// --- Siemens Structured Format ---
DATA_BLOCK "model__HS8_IW10_"
{ S7_Optimized_Access := 'TRUE' }
VERSION :
NON_RETAIN
   VAR
      W_i : ARRAY[0..7, 0..39] OF REAL;
      W_f : ARRAY[0..7, 0..39] OF REAL;
      W_g : ARRAY[0..7, 0..39] OF REAL;
      W_o : ARRAY[0..7, 0..39] OF REAL;
      R_i : ARRAY[0..7, 0..7] OF REAL;
      R_f : ARRAY[0..7, 0..7] OF REAL;
      R_g : ARRAY[0..7, 0..7] OF REAL;
      R_o : ARRAY[0..7, 0..7] OF REAL;
      B_i : ARRAY[0..7] OF REAL;
      B_f : ARRAY[0..7] OF REAL;
      B_g : ARRAY[0..7] OF REAL;
      B_o : ARRAY[0..7] OF REAL;
      FC_W : ARRAY[0..39, 0..7] OF REAL;
      FC_B : ARRAY[0..39] OF REAL;
   END_VAR
BEGIN

      W_i[0,0] := -0.07214709;
      W_i[0,1] := 0.05972328;
      W_i[0,2] := 0.02437277;
      W_i[0,3] := -0.07067372;
      W_i[0,4] := 0.15626091;
      W_i[0,5] := 0.03422371;
      W_i[0,6] := -0.01010964;
      W_i[0,7] := 0.24618091;
      W_i[0,8] := 0.19837169;
      W_i[0,9] := -0.16936609;
      W_i[0,10] := -0.03685989;
      W_i[0,11] := -0.34127542;
      W_i[0,12] := 0.16145179;
      W_i[0,13] := -0.03563828;
      W_i[0,14] := -0.03820900;
      W_i[0,15] := 0.03625023;
      W_i[0,16] := -0.00035658;
      W_i[0,17] := 0.05683306;
      W_i[0,18] := 0.01328012;
      W_i[0,19] := 0.01230632;
      W_i[0,20] := -0.02302203;
      W_i[0,21] := 0.29246566;
      W_i[0,22] := -0.40551317;
      W_i[0,23] := -0.00420093;
      W_i[0,24] := -0.49537772;
      W_i[0,25] := -0.37926760;
      W_i[0,26] := -0.32712772;
      W_i[0,27] := -0.47364110;
      W_i[0,28] := -0.02835605;
      W_i[0,29] := -0.19270489;
      W_i[0,30] := -0.02380528;
      W_i[0,31] := -0.25659311;
      W_i[0,32] := -0.07342248;
      W_i[0,33] := 0.12401358;
      W_i[0,34] := -0.00912032;
      W_i[0,35] := -0.27585000;
      W_i[0,36] := -0.01797117;
      W_i[0,37] := -0.35355157;
      W_i[0,38] := 0.03972119;
      W_i[0,39] := 0.01989586;
      W_i[1,0] := 0.10684982;
      W_i[1,1] := -0.11368593;
      W_i[1,2] := 0.13303033;
      W_i[1,3] := 0.06406520;
      W_i[1,4] := 0.10692474;
      W_i[1,5] := -0.00541547;
      W_i[1,6] := 0.13554892;
      W_i[1,7] := 0.02475992;
      W_i[1,8] := 0.05082010;
      W_i[1,9] := -0.42398453;
      W_i[1,10] := 0.03934563;
      W_i[1,11] := 0.28041703;
      W_i[1,12] := -0.48703033;
      W_i[1,13] := -0.03745792;
      W_i[1,14] := -0.00239940;
      W_i[1,15] := 0.15541774;
      W_i[1,16] := 0.04951616;
      W_i[1,17] := -0.01560813;
      W_i[1,18] := -0.00796859;
      W_i[1,19] := 0.12689193;
      W_i[1,20] := -0.06697816;
      W_i[1,21] := 0.18759193;
      W_i[1,22] := -0.37609926;
      W_i[1,23] := -0.01051652;
      W_i[1,24] := 0.38811579;
      W_i[1,25] := 0.20634656;
      W_i[1,26] := -0.03610945;
      W_i[1,27] := -0.06391723;
      W_i[1,28] := 0.06933470;
      W_i[1,29] := -0.03307433;
      W_i[1,30] := -0.16139032;
      W_i[1,31] := -0.13275333;
      W_i[1,32] := 0.16665860;
      W_i[1,33] := -0.25067136;
      W_i[1,34] := -0.03715657;
      W_i[1,35] := -0.52275580;
      W_i[1,36] := 0.03904245;
      W_i[1,37] := -0.14358856;
      W_i[1,38] := -0.15253240;
      W_i[1,39] := 0.02192211;
      W_i[2,0] := 0.00334517;
      W_i[2,1] := 0.09885125;
      W_i[2,2] := 0.04071221;
      W_i[2,3] := 0.04674324;
      W_i[2,4] := 0.04530917;
      W_i[2,5] := 0.10125730;
      W_i[2,6] := 0.06720760;
      W_i[2,7] := 0.00911526;
      W_i[2,8] := 0.07727423;
      W_i[2,9] := 0.03502122;
      W_i[2,10] := 0.02252782;
      W_i[2,11] := 0.14928287;
      W_i[2,12] := -0.06610898;
      W_i[2,13] := 0.07412212;
      W_i[2,14] := -0.01351282;
      W_i[2,15] := -0.06538101;
      W_i[2,16] := -0.05425974;
      W_i[2,17] := -0.05741069;
      W_i[2,18] := 0.50298566;
      W_i[2,19] := 0.05811854;
      W_i[2,20] := -0.03235166;
      W_i[2,21] := 0.02004486;
      W_i[2,22] := -0.02004233;
      W_i[2,23] := 0.00046481;
      W_i[2,24] := -0.34728089;
      W_i[2,25] := -0.59973961;
      W_i[2,26] := 0.09884801;
      W_i[2,27] := 0.08079667;
      W_i[2,28] := -0.06159005;
      W_i[2,29] := -0.21210669;
      W_i[2,30] := -0.02564744;
      W_i[2,31] := 0.03398452;
      W_i[2,32] := 0.07429420;
      W_i[2,33] := -0.16060953;
      W_i[2,34] := -0.61966300;
      W_i[2,35] := -0.02510496;
      W_i[2,36] := -0.09424359;
      W_i[2,37] := -0.20125464;
      W_i[2,38] := -0.02379467;
      W_i[2,39] := 0.00389740;
      W_i[3,0] := -0.41209814;
      W_i[3,1] := 0.07958311;
      W_i[3,2] := -0.04647379;
      W_i[3,3] := -0.35490474;
      W_i[3,4] := -0.16210698;
      W_i[3,5] := -0.05668240;
      W_i[3,6] := -0.06754937;
      W_i[3,7] := -0.41626674;
      W_i[3,8] := -0.45890990;
      W_i[3,9] := 0.37057030;
      W_i[3,10] := -0.02326192;
      W_i[3,11] := 0.25959259;
      W_i[3,12] := 0.01613945;
      W_i[3,13] := 0.14936726;
      W_i[3,14] := -0.02081729;
      W_i[3,15] := 0.03732191;
      W_i[3,16] := 0.01341023;
      W_i[3,17] := 0.04394821;
      W_i[3,18] := 0.13104227;
      W_i[3,19] := 0.08449978;
      W_i[3,20] := 0.16582783;
      W_i[3,21] := 0.00154001;
      W_i[3,22] := 0.15525876;
      W_i[3,23] := -0.21071896;
      W_i[3,24] := -0.06380144;
      W_i[3,25] := 0.10770430;
      W_i[3,26] := 0.13004155;
      W_i[3,27] := 0.18728302;
      W_i[3,28] := -0.45115548;
      W_i[3,29] := -0.00978980;
      W_i[3,30] := -0.01092611;
      W_i[3,31] := -0.13163096;
      W_i[3,32] := -0.06683033;
      W_i[3,33] := -0.17569157;
      W_i[3,34] := 0.41024187;
      W_i[3,35] := -0.29703203;
      W_i[3,36] := -0.00256490;
      W_i[3,37] := 0.07302216;
      W_i[3,38] := 0.19801962;
      W_i[3,39] := -0.14404945;
      W_i[4,0] := 0.00010722;
      W_i[4,1] := 0.05229621;
      W_i[4,2] := -0.05357129;
      W_i[4,3] := -0.14613566;
      W_i[4,4] := 0.00491695;
      W_i[4,5] := -0.01530431;
      W_i[4,6] := -0.07012728;
      W_i[4,7] := 0.12999427;
      W_i[4,8] := 0.01473324;
      W_i[4,9] := -0.13760696;
      W_i[4,10] := -0.07251389;
      W_i[4,11] := -0.00740168;
      W_i[4,12] := 0.04622447;
      W_i[4,13] := 0.03605191;
      W_i[4,14] := 0.02809449;
      W_i[4,15] := 0.03771993;
      W_i[4,16] := -0.01435529;
      W_i[4,17] := -0.03196694;
      W_i[4,18] := 0.09073107;
      W_i[4,19] := -0.04999484;
      W_i[4,20] := 0.05219137;
      W_i[4,21] := -0.08050881;
      W_i[4,22] := -0.04031698;
      W_i[4,23] := -0.13835990;
      W_i[4,24] := -0.43295500;
      W_i[4,25] := -0.05190322;
      W_i[4,26] := 0.17071831;
      W_i[4,27] := 0.03228986;
      W_i[4,28] := -0.04205497;
      W_i[4,29] := -0.08100788;
      W_i[4,30] := -0.15932465;
      W_i[4,31] := -0.13447607;
      W_i[4,32] := 0.12402157;
      W_i[4,33] := 0.18587913;
      W_i[4,34] := 0.31666172;
      W_i[4,35] := -0.12810661;
      W_i[4,36] := -0.01452139;
      W_i[4,37] := -0.07046619;
      W_i[4,38] := 0.03673343;
      W_i[4,39] := 0.10715080;
      W_i[5,0] := -0.13978986;
      W_i[5,1] := -0.07236300;
      W_i[5,2] := 0.01403345;
      W_i[5,3] := -0.08823197;
      W_i[5,4] := -0.11757445;
      W_i[5,5] := 0.03605668;
      W_i[5,6] := -0.00657548;
      W_i[5,7] := -0.41652936;
      W_i[5,8] := -0.16638683;
      W_i[5,9] := 0.44695261;
      W_i[5,10] := -0.02933357;
      W_i[5,11] := 0.13875259;
      W_i[5,12] := -0.00749722;
      W_i[5,13] := 0.00454487;
      W_i[5,14] := -0.00728751;
      W_i[5,15] := -0.05415151;
      W_i[5,16] := -0.00496033;
      W_i[5,17] := 0.01153068;
      W_i[5,18] := 0.11538580;
      W_i[5,19] := 0.04499825;
      W_i[5,20] := 0.06127532;
      W_i[5,21] := 0.06778700;
      W_i[5,22] := -0.34379280;
      W_i[5,23] := 0.14505032;
      W_i[5,24] := -0.56446981;
      W_i[5,25] := 0.02404343;
      W_i[5,26] := 0.06535989;
      W_i[5,27] := 0.06723037;
      W_i[5,28] := 0.08955745;
      W_i[5,29] := -0.00632868;
      W_i[5,30] := -0.47079688;
      W_i[5,31] := 0.11328098;
      W_i[5,32] := 0.16523570;
      W_i[5,33] := 0.04812213;
      W_i[5,34] := 0.10470282;
      W_i[5,35] := 0.05655447;
      W_i[5,36] := 0.04768148;
      W_i[5,37] := -0.27433640;
      W_i[5,38] := 0.09722462;
      W_i[5,39] := 0.04700476;
      W_i[6,0] := -0.11920829;
      W_i[6,1] := -0.26365072;
      W_i[6,2] := 0.06434898;
      W_i[6,3] := -0.50198841;
      W_i[6,4] := -0.02251296;
      W_i[6,5] := -0.05062700;
      W_i[6,6] := 0.20673671;
      W_i[6,7] := -0.23902187;
      W_i[6,8] := 0.24789530;
      W_i[6,9] := -0.12560840;
      W_i[6,10] := 0.35302734;
      W_i[6,11] := -0.56945974;
      W_i[6,12] := -0.63313663;
      W_i[6,13] := 0.11470533;
      W_i[6,14] := 0.04041832;
      W_i[6,15] := -0.32986644;
      W_i[6,16] := 0.26582161;
      W_i[6,17] := -0.39063680;
      W_i[6,18] := 0.32249957;
      W_i[6,19] := 0.20544839;
      W_i[6,20] := 0.10993068;
      W_i[6,21] := 0.06042655;
      W_i[6,22] := 0.34672299;
      W_i[6,23] := 0.11707149;
      W_i[6,24] := 0.80769390;
      W_i[6,25] := 1.00853431;
      W_i[6,26] := 0.16334604;
      W_i[6,27] := -0.07016917;
      W_i[6,28] := 0.09314778;
      W_i[6,29] := -0.14730705;
      W_i[6,30] := 0.22153552;
      W_i[6,31] := -0.13013706;
      W_i[6,32] := 0.27963796;
      W_i[6,33] := 0.31636471;
      W_i[6,34] := 1.01684213;
      W_i[6,35] := -0.21782602;
      W_i[6,36] := 0.00761380;
      W_i[6,37] := -0.16414484;
      W_i[6,38] := -0.44388211;
      W_i[6,39] := 0.70731664;
      W_i[7,0] := 0.08101967;
      W_i[7,1] := -0.06116093;
      W_i[7,2] := 0.09811447;
      W_i[7,3] := -0.27039346;
      W_i[7,4] := 0.22495940;
      W_i[7,5] := -0.05012152;
      W_i[7,6] := -0.09069129;
      W_i[7,7] := 0.12504753;
      W_i[7,8] := 0.15236920;
      W_i[7,9] := -0.16411021;
      W_i[7,10] := 0.01840155;
      W_i[7,11] := -0.24652572;
      W_i[7,12] := -0.09115234;
      W_i[7,13] := -0.09178895;
      W_i[7,14] := 0.03458378;
      W_i[7,15] := 0.11195860;
      W_i[7,16] := -0.03420459;
      W_i[7,17] := 0.01046852;
      W_i[7,18] := -0.00015169;
      W_i[7,19] := -0.00696717;
      W_i[7,20] := 0.18236621;
      W_i[7,21] := 0.18826969;
      W_i[7,22] := -0.02247082;
      W_i[7,23] := -0.04479990;
      W_i[7,24] := -0.28694034;
      W_i[7,25] := 0.29932031;
      W_i[7,26] := 0.10229074;
      W_i[7,27] := -0.33169511;
      W_i[7,28] := 0.07270649;
      W_i[7,29] := 0.22570691;
      W_i[7,30] := 0.42579922;
      W_i[7,31] := -0.02785212;
      W_i[7,32] := -0.23787680;
      W_i[7,33] := 0.30205894;
      W_i[7,34] := 0.48473808;
      W_i[7,35] := 0.03179261;
      W_i[7,36] := 0.02886904;
      W_i[7,37] := 0.21660374;
      W_i[7,38] := 0.05787315;
      W_i[7,39] := -0.04931584;
      W_f[0,0] := 0.00708323;
      W_f[0,1] := -0.01181322;
      W_f[0,2] := -0.11819337;
      W_f[0,3] := 0.13899828;
      W_f[0,4] := -0.02075264;
      W_f[0,5] := -0.03891272;
      W_f[0,6] := -0.07379504;
      W_f[0,7] := -0.11890592;
      W_f[0,8] := -0.09191579;
      W_f[0,9] := 0.12965402;
      W_f[0,10] := 0.02389325;
      W_f[0,11] := 0.05123832;
      W_f[0,12] := -0.18012317;
      W_f[0,13] := -0.05337619;
      W_f[0,14] := -0.07043158;
      W_f[0,15] := -0.11247810;
      W_f[0,16] := 0.09422214;
      W_f[0,17] := 0.21282011;
      W_f[0,18] := 0.05499737;
      W_f[0,19] := 0.10524461;
      W_f[0,20] := 0.06727590;
      W_f[0,21] := 0.18237843;
      W_f[0,22] := -0.02546566;
      W_f[0,23] := -0.06223162;
      W_f[0,24] := 0.71843404;
      W_f[0,25] := 0.81493032;
      W_f[0,26] := 0.03257482;
      W_f[0,27] := -0.07486192;
      W_f[0,28] := 0.04440695;
      W_f[0,29] := 0.17049384;
      W_f[0,30] := 0.15490918;
      W_f[0,31] := 0.10427933;
      W_f[0,32] := 0.13195500;
      W_f[0,33] := 0.02894589;
      W_f[0,34] := 0.95351958;
      W_f[0,35] := 0.13739404;
      W_f[0,36] := 0.03780418;
      W_f[0,37] := 0.12029935;
      W_f[0,38] := -0.13034570;
      W_f[0,39] := 0.17043786;
      W_f[1,0] := -0.05103588;
      W_f[1,1] := 0.03097129;
      W_f[1,2] := -0.03529896;
      W_f[1,3] := -0.08949374;
      W_f[1,4] := 0.05201217;
      W_f[1,5] := 0.07057156;
      W_f[1,6] := 0.04444524;
      W_f[1,7] := 0.13214116;
      W_f[1,8] := -0.18349366;
      W_f[1,9] := 0.09771031;
      W_f[1,10] := -0.02543963;
      W_f[1,11] := -0.15101723;
      W_f[1,12] := 0.09257572;
      W_f[1,13] := -0.02058279;
      W_f[1,14] := 0.04750511;
      W_f[1,15] := 0.00256356;
      W_f[1,16] := 0.03240434;
      W_f[1,17] := 0.02959783;
      W_f[1,18] := -0.07903013;
      W_f[1,19] := 0.06137549;
      W_f[1,20] := -0.08425386;
      W_f[1,21] := 0.04098953;
      W_f[1,22] := 0.37306514;
      W_f[1,23] := -0.01071887;
      W_f[1,24] := 0.89733803;
      W_f[1,25] := 1.21406257;
      W_f[1,26] := 0.06516311;
      W_f[1,27] := 0.00914704;
      W_f[1,28] := 0.04227815;
      W_f[1,29] := -0.10532902;
      W_f[1,30] := 0.16040285;
      W_f[1,31] := -0.10591315;
      W_f[1,32] := 0.31760797;
      W_f[1,33] := 0.05462405;
      W_f[1,34] := 1.00453556;
      W_f[1,35] := -0.27051091;
      W_f[1,36] := -0.05915660;
      W_f[1,37] := 0.28985777;
      W_f[1,38] := -0.00542082;
      W_f[1,39] := 0.24056318;
      W_f[2,0] := 0.12671420;
      W_f[2,1] := -0.10912015;
      W_f[2,2] := 0.09372077;
      W_f[2,3] := -0.06474926;
      W_f[2,4] := -0.21063805;
      W_f[2,5] := -0.02976029;
      W_f[2,6] := -0.03741420;
      W_f[2,7] := -0.02389968;
      W_f[2,8] := -0.10062340;
      W_f[2,9] := -0.03533751;
      W_f[2,10] := -0.03556222;
      W_f[2,11] := -0.18180723;
      W_f[2,12] := 0.00197740;
      W_f[2,13] := 0.13552259;
      W_f[2,14] := -0.01979193;
      W_f[2,15] := 0.02504811;
      W_f[2,16] := -0.00935277;
      W_f[2,17] := -0.00082860;
      W_f[2,18] := 0.02693685;
      W_f[2,19] := -0.09008320;
      W_f[2,20] := -0.02276102;
      W_f[2,21] := -0.03999444;
      W_f[2,22] := -0.02197137;
      W_f[2,23] := 0.23856066;
      W_f[2,24] := 0.09475329;
      W_f[2,25] := -0.13239257;
      W_f[2,26] := -0.02748259;
      W_f[2,27] := -0.16801514;
      W_f[2,28] := 0.02366016;
      W_f[2,29] := 0.37193993;
      W_f[2,30] := -0.03538382;
      W_f[2,31] := 0.00506000;
      W_f[2,32] := -0.12670894;
      W_f[2,33] := 0.20883897;
      W_f[2,34] := -0.46258271;
      W_f[2,35] := 0.32857734;
      W_f[2,36] := 0.03205189;
      W_f[2,37] := 0.06433915;
      W_f[2,38] := -0.00436854;
      W_f[2,39] := -0.04177000;
      W_f[3,0] := 0.09149595;
      W_f[3,1] := 0.05684213;
      W_f[3,2] := -0.04046491;
      W_f[3,3] := 0.16697308;
      W_f[3,4] := -0.24152677;
      W_f[3,5] := -0.04763369;
      W_f[3,6] := -0.21290614;
      W_f[3,7] := 0.17224246;
      W_f[3,8] := -0.02882880;
      W_f[3,9] := -0.34723446;
      W_f[3,10] := 0.13916484;
      W_f[3,11] := -0.17330380;
      W_f[3,12] := -0.07241807;
      W_f[3,13] := -0.18257356;
      W_f[3,14] := -0.07163820;
      W_f[3,15] := 0.13798824;
      W_f[3,16] := 0.03025815;
      W_f[3,17] := 0.13978501;
      W_f[3,18] := -1.50750315;
      W_f[3,19] := 0.05514524;
      W_f[3,20] := -0.02955024;
      W_f[3,21] := -0.08395630;
      W_f[3,22] := -0.16754888;
      W_f[3,23] := 0.01334867;
      W_f[3,24] := -0.07160708;
      W_f[3,25] := -0.32795355;
      W_f[3,26] := -0.43044916;
      W_f[3,27] := 0.05751909;
      W_f[3,28] := 0.06252181;
      W_f[3,29] := 0.50739962;
      W_f[3,30] := -0.00872058;
      W_f[3,31] := 0.13262282;
      W_f[3,32] := 0.40081328;
      W_f[3,33] := 0.06643189;
      W_f[3,34] := -0.29172045;
      W_f[3,35] := 0.30180812;
      W_f[3,36] := 0.11044914;
      W_f[3,37] := -0.04694669;
      W_f[3,38] := -0.00254733;
      W_f[3,39] := -0.10670592;
      W_f[4,0] := -0.04173987;
      W_f[4,1] := -0.00443699;
      W_f[4,2] := -0.01804712;
      W_f[4,3] := 0.02465925;
      W_f[4,4] := 0.10097732;
      W_f[4,5] := 0.00270554;
      W_f[4,6] := -0.00317248;
      W_f[4,7] := -0.18945615;
      W_f[4,8] := -0.10332906;
      W_f[4,9] := 0.05336653;
      W_f[4,10] := 0.01227043;
      W_f[4,11] := -0.02219165;
      W_f[4,12] := -0.03810129;
      W_f[4,13] := -0.03208273;
      W_f[4,14] := 0.04131512;
      W_f[4,15] := -0.03503123;
      W_f[4,16] := 0.04256575;
      W_f[4,17] := -0.03164240;
      W_f[4,18] := 0.04763466;
      W_f[4,19] := 0.04308751;
      W_f[4,20] := 0.06900967;
      W_f[4,21] := -0.08195710;
      W_f[4,22] := 0.11304240;
      W_f[4,23] := 0.09688803;
      W_f[4,24] := -0.50463659;
      W_f[4,25] := -0.38656512;
      W_f[4,26] := -0.13179161;
      W_f[4,27] := 0.01542916;
      W_f[4,28] := 0.07802795;
      W_f[4,29] := -0.14032713;
      W_f[4,30] := 0.14824803;
      W_f[4,31] := 0.12095391;
      W_f[4,32] := 0.02171578;
      W_f[4,33] := -0.15110554;
      W_f[4,34] := -0.18883832;
      W_f[4,35] := -0.03473442;
      W_f[4,36] := 0.05890166;
      W_f[4,37] := -0.01619323;
      W_f[4,38] := 0.04949700;
      W_f[4,39] := 0.07575098;
      W_f[5,0] := -0.09567674;
      W_f[5,1] := 0.09717870;
      W_f[5,2] := 0.03514667;
      W_f[5,3] := 0.05669624;
      W_f[5,4] := -0.02355025;
      W_f[5,5] := -0.00160842;
      W_f[5,6] := 0.09726227;
      W_f[5,7] := -0.43277800;
      W_f[5,8] := -0.15966371;
      W_f[5,9] := 0.38071355;
      W_f[5,10] := 0.00158656;
      W_f[5,11] := 0.17037611;
      W_f[5,12] := -0.08529956;
      W_f[5,13] := 0.00575568;
      W_f[5,14] := 0.07765908;
      W_f[5,15] := -0.13563958;
      W_f[5,16] := -0.10357573;
      W_f[5,17] := -0.20172329;
      W_f[5,18] := -0.13053854;
      W_f[5,19] := 0.03271331;
      W_f[5,20] := -0.03536206;
      W_f[5,21] := 0.14749785;
      W_f[5,22] := 0.46310273;
      W_f[5,23] := -0.03476221;
      W_f[5,24] := 1.87947142;
      W_f[5,25] := 1.58035707;
      W_f[5,26] := -0.05445153;
      W_f[5,27] := -0.16590932;
      W_f[5,28] := 0.10555614;
      W_f[5,29] := -0.22020321;
      W_f[5,30] := 0.59286916;
      W_f[5,31] := 0.05095429;
      W_f[5,32] := 0.19744034;
      W_f[5,33] := 0.25974834;
      W_f[5,34] := 1.41725945;
      W_f[5,35] := -0.05630583;
      W_f[5,36] := -0.00765480;
      W_f[5,37] := 0.11030062;
      W_f[5,38] := 0.07699158;
      W_f[5,39] := 0.51856029;
      W_f[6,0] := 0.04847221;
      W_f[6,1] := 0.04356489;
      W_f[6,2] := -0.04560984;
      W_f[6,3] := 0.04543123;
      W_f[6,4] := 0.04954825;
      W_f[6,5] := 0.00071875;
      W_f[6,6] := -0.07963482;
      W_f[6,7] := 0.04270557;
      W_f[6,8] := -0.06502789;
      W_f[6,9] := -0.13146918;
      W_f[6,10] := -0.07300840;
      W_f[6,11] := -0.06714232;
      W_f[6,12] := 0.18289082;
      W_f[6,13] := -0.04542018;
      W_f[6,14] := -0.00317417;
      W_f[6,15] := -0.00539382;
      W_f[6,16] := 0.00731518;
      W_f[6,17] := -0.09440549;
      W_f[6,18] := -0.06629226;
      W_f[6,19] := -0.10041165;
      W_f[6,20] := 0.06385964;
      W_f[6,21] := -0.00066353;
      W_f[6,22] := 0.11827765;
      W_f[6,23] := -0.01271241;
      W_f[6,24] := 1.09554279;
      W_f[6,25] := 1.13105202;
      W_f[6,26] := 0.06568716;
      W_f[6,27] := -0.03536376;
      W_f[6,28] := 0.02383021;
      W_f[6,29] := 0.05406570;
      W_f[6,30] := 0.15167096;
      W_f[6,31] := -0.02357897;
      W_f[6,32] := 0.03374309;
      W_f[6,33] := 0.14940892;
      W_f[6,34] := 0.85827291;
      W_f[6,35] := 0.10391039;
      W_f[6,36] := -0.01731022;
      W_f[6,37] := -0.01241286;
      W_f[6,38] := -0.07383022;
      W_f[6,39] := 0.23319298;
      W_f[7,0] := -0.00703594;
      W_f[7,1] := 0.01558984;
      W_f[7,2] := -0.00251701;
      W_f[7,3] := 0.14500660;
      W_f[7,4] := 0.05646368;
      W_f[7,5] := -0.01658792;
      W_f[7,6] := -0.09505704;
      W_f[7,7] := 0.02159695;
      W_f[7,8] := -0.16402565;
      W_f[7,9] := 0.00675202;
      W_f[7,10] := -0.05481035;
      W_f[7,11] := -0.13274667;
      W_f[7,12] := 0.24241473;
      W_f[7,13] := 0.00729740;
      W_f[7,14] := -0.14640833;
      W_f[7,15] := -0.04770046;
      W_f[7,16] := 0.14853485;
      W_f[7,17] := 0.00505042;
      W_f[7,18] := -0.00851168;
      W_f[7,19] := -0.20896289;
      W_f[7,20] := 0.02721659;
      W_f[7,21] := 0.08800104;
      W_f[7,22] := 0.06278189;
      W_f[7,23] := -0.00083155;
      W_f[7,24] := 1.37909341;
      W_f[7,25] := 1.16676664;
      W_f[7,26] := -0.00847061;
      W_f[7,27] := -0.02336962;
      W_f[7,28] := 0.00882273;
      W_f[7,29] := 0.35906574;
      W_f[7,30] := 0.08403210;
      W_f[7,31] := -0.03630471;
      W_f[7,32] := 0.19077916;
      W_f[7,33] := 0.20514297;
      W_f[7,34] := 0.21810204;
      W_f[7,35] := 0.06294452;
      W_f[7,36] := 0.00392204;
      W_f[7,37] := 0.09456417;
      W_f[7,38] := -0.01927309;
      W_f[7,39] := 0.27183673;
      W_g[0,0] := -0.07034334;
      W_g[0,1] := 0.03156179;
      W_g[0,2] := -0.06465199;
      W_g[0,3] := 0.01206673;
      W_g[0,4] := -0.11430016;
      W_g[0,5] := -0.01664878;
      W_g[0,6] := 0.02142663;
      W_g[0,7] := 0.01663074;
      W_g[0,8] := 0.02022547;
      W_g[0,9] := 0.01864452;
      W_g[0,10] := 0.00190711;
      W_g[0,11] := 0.00721099;
      W_g[0,12] := 0.02579849;
      W_g[0,13] := -0.03713468;
      W_g[0,14] := -0.06940822;
      W_g[0,15] := -0.01003235;
      W_g[0,16] := 0.00773649;
      W_g[0,17] := 0.11996724;
      W_g[0,18] := 0.02323754;
      W_g[0,19] := 0.00800148;
      W_g[0,20] := -0.02301983;
      W_g[0,21] := 0.10161702;
      W_g[0,22] := 0.03288819;
      W_g[0,23] := -0.03117830;
      W_g[0,24] := 0.48237947;
      W_g[0,25] := 0.36674199;
      W_g[0,26] := -0.05521943;
      W_g[0,27] := 0.12540811;
      W_g[0,28] := -0.12757246;
      W_g[0,29] := -0.03407666;
      W_g[0,30] := 0.01104811;
      W_g[0,31] := 0.02846052;
      W_g[0,32] := 0.00676780;
      W_g[0,33] := 0.02226435;
      W_g[0,34] := -0.05392364;
      W_g[0,35] := 0.01852163;
      W_g[0,36] := 0.07350205;
      W_g[0,37] := 0.05389259;
      W_g[0,38] := -0.05447108;
      W_g[0,39] := -0.07045685;
      W_g[1,0] := -0.00444380;
      W_g[1,1] := 0.00524623;
      W_g[1,2] := -0.00320254;
      W_g[1,3] := 0.01111780;
      W_g[1,4] := -0.02181038;
      W_g[1,5] := -0.06435853;
      W_g[1,6] := -0.11283723;
      W_g[1,7] := 0.00893267;
      W_g[1,8] := 0.01303838;
      W_g[1,9] := 0.00185226;
      W_g[1,10] := 0.06878208;
      W_g[1,11] := 0.07648126;
      W_g[1,12] := 0.07980552;
      W_g[1,13] := 0.01262750;
      W_g[1,14] := -0.03160430;
      W_g[1,15] := 0.10011385;
      W_g[1,16] := -0.09624640;
      W_g[1,17] := -0.12084271;
      W_g[1,18] := -0.02024449;
      W_g[1,19] := 0.07013080;
      W_g[1,20] := 0.10538352;
      W_g[1,21] := -0.03829639;
      W_g[1,22] := -0.00354391;
      W_g[1,23] := 0.03275719;
      W_g[1,24] := 0.17965782;
      W_g[1,25] := -0.19564816;
      W_g[1,26] := 0.00854688;
      W_g[1,27] := -0.03361512;
      W_g[1,28] := -0.07664448;
      W_g[1,29] := -0.00350407;
      W_g[1,30] := 0.00330394;
      W_g[1,31] := 0.00362330;
      W_g[1,32] := -0.00242198;
      W_g[1,33] := 0.00457848;
      W_g[1,34] := 0.41679174;
      W_g[1,35] := 0.03201690;
      W_g[1,36] := 0.01899636;
      W_g[1,37] := -0.04047984;
      W_g[1,38] := -0.05404723;
      W_g[1,39] := -0.03850636;
      W_g[2,0] := 0.09367149;
      W_g[2,1] := 0.00112518;
      W_g[2,2] := 0.08251125;
      W_g[2,3] := -0.01032626;
      W_g[2,4] := -0.17358032;
      W_g[2,5] := 0.06058484;
      W_g[2,6] := 0.04647175;
      W_g[2,7] := -0.01058286;
      W_g[2,8] := -0.00198453;
      W_g[2,9] := -0.00400265;
      W_g[2,10] := -0.00210860;
      W_g[2,11] := -0.05763165;
      W_g[2,12] := -0.02976729;
      W_g[2,13] := 0.16225053;
      W_g[2,14] := -0.01911786;
      W_g[2,15] := -0.02073957;
      W_g[2,16] := -0.02424970;
      W_g[2,17] := -0.02491161;
      W_g[2,18] := -0.14540172;
      W_g[2,19] := 0.01427219;
      W_g[2,20] := -0.05718472;
      W_g[2,21] := -0.00834007;
      W_g[2,22] := 0.01367352;
      W_g[2,23] := 0.16430169;
      W_g[2,24] := 0.32054973;
      W_g[2,25] := 0.38814557;
      W_g[2,26] := 0.07002852;
      W_g[2,27] := 0.02144061;
      W_g[2,28] := -0.07323609;
      W_g[2,29] := 0.01338264;
      W_g[2,30] := 0.02144418;
      W_g[2,31] := 0.01571183;
      W_g[2,32] := 0.01401756;
      W_g[2,33] := 0.00919776;
      W_g[2,34] := 0.87235081;
      W_g[2,35] := -0.07491063;
      W_g[2,36] := -0.04177252;
      W_g[2,37] := 0.09778510;
      W_g[2,38] := -0.02624917;
      W_g[2,39] := -0.01247705;
      W_g[3,0] := -0.00312740;
      W_g[3,1] := 0.01748835;
      W_g[3,2] := -0.00530153;
      W_g[3,3] := -0.03639691;
      W_g[3,4] := -0.09401610;
      W_g[3,5] := -0.02446339;
      W_g[3,6] := -0.05136326;
      W_g[3,7] := -0.02695942;
      W_g[3,8] := -0.02937514;
      W_g[3,9] := -0.03799582;
      W_g[3,10] := 0.00379267;
      W_g[3,11] := -0.03588169;
      W_g[3,12] := -0.02958600;
      W_g[3,13] := 0.01290534;
      W_g[3,14] := 0.02873308;
      W_g[3,15] := -0.02114533;
      W_g[3,16] := 0.00849492;
      W_g[3,17] := -0.02519036;
      W_g[3,18] := -0.11424359;
      W_g[3,19] := -0.03385856;
      W_g[3,20] := 0.03059323;
      W_g[3,21] := 0.01884498;
      W_g[3,22] := -0.03800057;
      W_g[3,23] := 0.01210539;
      W_g[3,24] := -0.49563253;
      W_g[3,25] := -0.65994966;
      W_g[3,26] := -0.03385233;
      W_g[3,27] := 0.03389804;
      W_g[3,28] := -0.11069407;
      W_g[3,29] := 0.07897274;
      W_g[3,30] := -0.05612407;
      W_g[3,31] := -0.01165623;
      W_g[3,32] := -0.03924601;
      W_g[3,33] := -0.02041759;
      W_g[3,34] := -0.12063195;
      W_g[3,35] := -0.06332459;
      W_g[3,36] := 0.01482042;
      W_g[3,37] := 0.03349160;
      W_g[3,38] := 0.02928583;
      W_g[3,39] := 0.60842210;
      W_g[4,0] := 0.02868404;
      W_g[4,1] := -0.04825799;
      W_g[4,2] := 0.02482833;
      W_g[4,3] := 0.06132923;
      W_g[4,4] := -0.08855467;
      W_g[4,5] := 0.04589472;
      W_g[4,6] := 0.08157697;
      W_g[4,7] := 0.07234233;
      W_g[4,8] := 0.05229455;
      W_g[4,9] := 0.05496285;
      W_g[4,10] := 0.02096794;
      W_g[4,11] := 0.02207873;
      W_g[4,12] := 0.03108713;
      W_g[4,13] := 0.00665728;
      W_g[4,14] := -0.04965325;
      W_g[4,15] := 0.01889800;
      W_g[4,16] := -0.02251282;
      W_g[4,17] := 0.03557793;
      W_g[4,18] := -0.07591323;
      W_g[4,19] := 0.04966724;
      W_g[4,20] := -0.08873382;
      W_g[4,21] := 0.01310619;
      W_g[4,22] := -0.04439254;
      W_g[4,23] := 0.03415269;
      W_g[4,24] := -0.62770677;
      W_g[4,25] := -0.10581250;
      W_g[4,26] := -0.01891168;
      W_g[4,27] := 0.02480597;
      W_g[4,28] := -0.00201301;
      W_g[4,29] := 0.07145379;
      W_g[4,30] := -0.04382761;
      W_g[4,31] := -0.04298389;
      W_g[4,32] := -0.02887516;
      W_g[4,33] := -0.03160532;
      W_g[4,34] := 0.21834604;
      W_g[4,35] := 0.01873893;
      W_g[4,36] := -0.06442018;
      W_g[4,37] := -0.11304606;
      W_g[4,38] := -0.04509857;
      W_g[4,39] := -0.02925531;
      W_g[5,0] := 0.18268949;
      W_g[5,1] := -0.11797520;
      W_g[5,2] := 0.17629275;
      W_g[5,3] := 0.03142028;
      W_g[5,4] := -0.01652149;
      W_g[5,5] := -0.05967048;
      W_g[5,6] := -0.04142075;
      W_g[5,7] := 0.02769361;
      W_g[5,8] := 0.02803064;
      W_g[5,9] := 0.04083285;
      W_g[5,10] := 0.03677053;
      W_g[5,11] := -0.07351185;
      W_g[5,12] := -0.08407787;
      W_g[5,13] := 0.03595718;
      W_g[5,14] := -0.00242524;
      W_g[5,15] := -0.06877073;
      W_g[5,16] := 0.00374599;
      W_g[5,17] := -0.03411847;
      W_g[5,18] := 0.06481477;
      W_g[5,19] := -0.09435212;
      W_g[5,20] := 0.04101316;
      W_g[5,21] := 0.04863375;
      W_g[5,22] := -0.02486804;
      W_g[5,23] := 0.04388688;
      W_g[5,24] := -0.10377861;
      W_g[5,25] := 0.35907325;
      W_g[5,26] := -0.04512582;
      W_g[5,27] := 0.06372260;
      W_g[5,28] := -0.04580466;
      W_g[5,29] := 0.00918311;
      W_g[5,30] := -0.05401663;
      W_g[5,31] := 0.01057453;
      W_g[5,32] := -0.04817041;
      W_g[5,33] := -0.03328571;
      W_g[5,34] := -0.01978806;
      W_g[5,35] := -0.08799826;
      W_g[5,36] := 0.06790313;
      W_g[5,37] := 0.09022456;
      W_g[5,38] := 0.01308107;
      W_g[5,39] := 0.01720484;
      W_g[6,0] := 0.06210544;
      W_g[6,1] := -0.00964019;
      W_g[6,2] := 0.06184339;
      W_g[6,3] := -0.06458558;
      W_g[6,4] := -0.00151253;
      W_g[6,5] := 0.04355884;
      W_g[6,6] := 0.05581776;
      W_g[6,7] := -0.07905485;
      W_g[6,8] := -0.06635278;
      W_g[6,9] := -0.06286671;
      W_g[6,10] := -0.08623632;
      W_g[6,11] := -0.01245475;
      W_g[6,12] := -0.03378635;
      W_g[6,13] := 0.03127304;
      W_g[6,14] := -0.02078948;
      W_g[6,15] := 0.00137005;
      W_g[6,16] := -0.07733220;
      W_g[6,17] := -0.10649602;
      W_g[6,18] := 0.02146085;
      W_g[6,19] := -0.03412123;
      W_g[6,20] := -0.05842118;
      W_g[6,21] := 0.03570734;
      W_g[6,22] := -0.00927513;
      W_g[6,23] := -0.00962296;
      W_g[6,24] := 0.01154771;
      W_g[6,25] := 0.06284481;
      W_g[6,26] := -0.02478036;
      W_g[6,27] := 0.03437400;
      W_g[6,28] := 0.05358073;
      W_g[6,29] := 0.01064103;
      W_g[6,30] := -0.00959687;
      W_g[6,31] := -0.00935796;
      W_g[6,32] := -0.01104967;
      W_g[6,33] := -0.00710198;
      W_g[6,34] := 0.27764010;
      W_g[6,35] := -0.04841734;
      W_g[6,36] := 0.00098623;
      W_g[6,37] := 0.03043675;
      W_g[6,38] := -0.03496779;
      W_g[6,39] := -0.02783902;
      W_g[7,0] := 0.03619956;
      W_g[7,1] := -0.01139570;
      W_g[7,2] := 0.03186626;
      W_g[7,3] := -0.02594865;
      W_g[7,4] := 0.11965120;
      W_g[7,5] := -0.03254651;
      W_g[7,6] := -0.07578963;
      W_g[7,7] := -0.03363758;
      W_g[7,8] := -0.03082440;
      W_g[7,9] := -0.02712537;
      W_g[7,10] := 0.00642671;
      W_g[7,11] := -0.08782534;
      W_g[7,12] := -0.09268230;
      W_g[7,13] := 0.00914687;
      W_g[7,14] := -0.08760387;
      W_g[7,15] := -0.11542334;
      W_g[7,16] := 0.00707082;
      W_g[7,17] := 0.11704925;
      W_g[7,18] := 0.05226066;
      W_g[7,19] := -0.08682797;
      W_g[7,20] := 0.07598362;
      W_g[7,21] := -0.08286781;
      W_g[7,22] := -0.01627091;
      W_g[7,23] := -0.01264957;
      W_g[7,24] := -0.47079486;
      W_g[7,25] := -0.07540244;
      W_g[7,26] := 0.02426168;
      W_g[7,27] := -0.07233322;
      W_g[7,28] := 0.05062053;
      W_g[7,29] := 0.02186041;
      W_g[7,30] := -0.01840415;
      W_g[7,31] := -0.00962791;
      W_g[7,32] := -0.02041369;
      W_g[7,33] := -0.02006152;
      W_g[7,34] := -0.07425848;
      W_g[7,35] := -0.06536297;
      W_g[7,36] := -0.00430546;
      W_g[7,37] := 0.04031537;
      W_g[7,38] := -0.06503575;
      W_g[7,39] := -0.08399117;
      W_o[0,0] := -0.57085669;
      W_o[0,1] := -0.04681201;
      W_o[0,2] := -0.24800207;
      W_o[0,3] := -0.38602149;
      W_o[0,4] := -0.34429318;
      W_o[0,5] := 0.10549517;
      W_o[0,6] := -0.26367727;
      W_o[0,7] := -0.13702963;
      W_o[0,8] := -0.15231206;
      W_o[0,9] := -0.14323375;
      W_o[0,10] := -0.13618764;
      W_o[0,11] := 0.08623260;
      W_o[0,12] := 0.20636982;
      W_o[0,13] := -0.03830929;
      W_o[0,14] := 0.12331601;
      W_o[0,15] := 0.02166978;
      W_o[0,16] := -0.08123493;
      W_o[0,17] := -0.08618607;
      W_o[0,18] := 0.54233044;
      W_o[0,19] := -0.11915454;
      W_o[0,20] := -0.32456002;
      W_o[0,21] := -0.03020910;
      W_o[0,22] := 0.65767694;
      W_o[0,23] := -0.04952972;
      W_o[0,24] := 1.36234951;
      W_o[0,25] := 1.66532695;
      W_o[0,26] := -0.74773312;
      W_o[0,27] := 0.15801664;
      W_o[0,28] := -0.01813998;
      W_o[0,29] := 0.02730388;
      W_o[0,30] := 0.43068638;
      W_o[0,31] := 0.36317101;
      W_o[0,32] := 0.06420399;
      W_o[0,33] := -0.20908703;
      W_o[0,34] := 1.31859016;
      W_o[0,35] := -0.21934026;
      W_o[0,36] := 0.26863953;
      W_o[0,37] := -0.11312449;
      W_o[0,38] := -0.11992589;
      W_o[0,39] := 0.99821264;
      W_o[1,0] := 0.10667461;
      W_o[1,1] := 0.01962533;
      W_o[1,2] := -0.00480660;
      W_o[1,3] := -0.00752457;
      W_o[1,4] := -0.11217720;
      W_o[1,5] := 0.00206603;
      W_o[1,6] := -0.07063800;
      W_o[1,7] := -0.08116529;
      W_o[1,8] := 0.04971202;
      W_o[1,9] := -0.02052844;
      W_o[1,10] := 0.06039909;
      W_o[1,11] := -0.32314682;
      W_o[1,12] := -0.11838520;
      W_o[1,13] := 0.04847965;
      W_o[1,14] := 0.01095985;
      W_o[1,15] := -0.07885160;
      W_o[1,16] := 0.22081691;
      W_o[1,17] := -0.01069563;
      W_o[1,18] := 0.05992901;
      W_o[1,19] := -0.02966248;
      W_o[1,20] := 0.43488529;
      W_o[1,21] := 0.06811651;
      W_o[1,22] := 0.06945629;
      W_o[1,23] := -0.06210565;
      W_o[1,24] := 1.04133368;
      W_o[1,25] := 0.79160953;
      W_o[1,26] := 0.15757442;
      W_o[1,27] := -0.09610198;
      W_o[1,28] := -0.15777384;
      W_o[1,29] := -0.26314041;
      W_o[1,30] := 0.22122788;
      W_o[1,31] := 0.01242414;
      W_o[1,32] := 0.11826468;
      W_o[1,33] := 0.09161918;
      W_o[1,34] := 0.96783555;
      W_o[1,35] := 0.08615178;
      W_o[1,36] := -0.06596540;
      W_o[1,37] := -0.20505081;
      W_o[1,38] := -0.12099239;
      W_o[1,39] := 0.81992567;
      W_o[2,0] := 0.07692418;
      W_o[2,1] := -0.11036226;
      W_o[2,2] := 0.02623424;
      W_o[2,3] := 0.02940779;
      W_o[2,4] := 0.08105131;
      W_o[2,5] := -0.07215023;
      W_o[2,6] := 0.05821245;
      W_o[2,7] := 0.12392700;
      W_o[2,8] := 0.00331179;
      W_o[2,9] := -0.20764571;
      W_o[2,10] := 0.32663119;
      W_o[2,11] := 0.02233894;
      W_o[2,12] := 0.07203373;
      W_o[2,13] := -0.37837738;
      W_o[2,14] := 0.15081947;
      W_o[2,15] := -0.04852225;
      W_o[2,16] := -0.06858451;
      W_o[2,17] := -0.04667585;
      W_o[2,18] := 1.27405727;
      W_o[2,19] := -0.02571864;
      W_o[2,20] := -0.01813021;
      W_o[2,21] := 0.68052500;
      W_o[2,22] := 0.22743875;
      W_o[2,23] := -0.67374688;
      W_o[2,24] := -0.30051517;
      W_o[2,25] := 0.09985244;
      W_o[2,26] := 0.01096807;
      W_o[2,27] := -0.04011973;
      W_o[2,28] := 0.36460930;
      W_o[2,29] := -0.13026837;
      W_o[2,30] := 0.17856032;
      W_o[2,31] := 0.14580105;
      W_o[2,32] := -0.01857202;
      W_o[2,33] := 0.36115634;
      W_o[2,34] := 0.18000041;
      W_o[2,35] := -0.01968618;
      W_o[2,36] := -0.11631926;
      W_o[2,37] := -0.22437349;
      W_o[2,38] := 0.36917746;
      W_o[2,39] := 0.18247823;
      W_o[3,0] := -0.25305161;
      W_o[3,1] := -0.05748865;
      W_o[3,2] := -0.14973676;
      W_o[3,3] := -0.34950122;
      W_o[3,4] := 0.17906217;
      W_o[3,5] := 0.33135971;
      W_o[3,6] := 0.54163671;
      W_o[3,7] := 0.18129022;
      W_o[3,8] := -0.21506567;
      W_o[3,9] := -0.16582678;
      W_o[3,10] := 0.03354707;
      W_o[3,11] := 0.03781534;
      W_o[3,12] := -0.74912232;
      W_o[3,13] := -0.00002978;
      W_o[3,14] := 0.10795104;
      W_o[3,15] := -0.00511314;
      W_o[3,16] := -0.00772868;
      W_o[3,17] := 0.11671072;
      W_o[3,18] := -0.05170535;
      W_o[3,19] := 0.01881175;
      W_o[3,20] := -0.05257827;
      W_o[3,21] := -0.00041528;
      W_o[3,22] := -0.11215112;
      W_o[3,23] := 0.03263832;
      W_o[3,24] := -0.49468938;
      W_o[3,25] := -0.16897368;
      W_o[3,26] := -0.00836590;
      W_o[3,27] := -0.12664883;
      W_o[3,28] := 0.41327897;
      W_o[3,29] := 0.15271561;
      W_o[3,30] := -0.00538531;
      W_o[3,31] := -0.19345705;
      W_o[3,32] := -0.13221580;
      W_o[3,33] := 0.35120431;
      W_o[3,34] := 0.06960481;
      W_o[3,35] := -0.06442323;
      W_o[3,36] := -0.17462859;
      W_o[3,37] := 0.00698183;
      W_o[3,38] := -0.11534231;
      W_o[3,39] := 0.12678961;
      W_o[4,0] := 0.30061489;
      W_o[4,1] := 0.29126322;
      W_o[4,2] := 0.01201630;
      W_o[4,3] := 0.11307906;
      W_o[4,4] := 0.05800173;
      W_o[4,5] := 0.05204230;
      W_o[4,6] := 0.14197972;
      W_o[4,7] := 0.35224134;
      W_o[4,8] := -0.06268087;
      W_o[4,9] := 0.33943415;
      W_o[4,10] := 0.05441138;
      W_o[4,11] := 0.03230330;
      W_o[4,12] := -0.11484767;
      W_o[4,13] := -0.08048104;
      W_o[4,14] := 0.04593046;
      W_o[4,15] := -0.12167345;
      W_o[4,16] := 0.01774614;
      W_o[4,17] := -0.06578777;
      W_o[4,18] := -0.21332319;
      W_o[4,19] := -0.25459981;
      W_o[4,20] := -0.15229602;
      W_o[4,21] := 0.18717009;
      W_o[4,22] := 0.04886236;
      W_o[4,23] := -0.03599270;
      W_o[4,24] := -0.04652552;
      W_o[4,25] := -0.24323644;
      W_o[4,26] := -0.17948933;
      W_o[4,27] := -0.25262487;
      W_o[4,28] := -0.15929545;
      W_o[4,29] := 0.04956881;
      W_o[4,30] := -0.28498772;
      W_o[4,31] := -0.10077197;
      W_o[4,32] := 0.07382053;
      W_o[4,33] := 0.04429949;
      W_o[4,34] := -0.05270445;
      W_o[4,35] := 0.13536042;
      W_o[4,36] := -0.01786239;
      W_o[4,37] := 0.31803700;
      W_o[4,38] := -0.13451934;
      W_o[4,39] := 0.56871533;
      W_o[5,0] := 0.38830724;
      W_o[5,1] := -0.67464000;
      W_o[5,2] := -0.03622986;
      W_o[5,3] := -0.31041449;
      W_o[5,4] := 0.03742103;
      W_o[5,5] := -0.06870902;
      W_o[5,6] := -0.17940173;
      W_o[5,7] := 0.16546406;
      W_o[5,8] := -0.50603092;
      W_o[5,9] := -0.10525495;
      W_o[5,10] := -0.32540444;
      W_o[5,11] := -0.31151175;
      W_o[5,12] := -0.20012428;
      W_o[5,13] := -0.24050371;
      W_o[5,14] := -0.12048050;
      W_o[5,15] := -0.38477761;
      W_o[5,16] := 0.14707315;
      W_o[5,17] := 0.47272572;
      W_o[5,18] := 0.35924280;
      W_o[5,19] := -0.34276947;
      W_o[5,20] := -0.09197704;
      W_o[5,21] := -0.11951853;
      W_o[5,22] := 0.13050619;
      W_o[5,23] := -0.37483913;
      W_o[5,24] := 2.15172362;
      W_o[5,25] := 1.96999085;
      W_o[5,26] := -0.56420952;
      W_o[5,27] := 0.07533623;
      W_o[5,28] := -0.22395705;
      W_o[5,29] := -0.10359064;
      W_o[5,30] := 0.33768624;
      W_o[5,31] := 0.01281008;
      W_o[5,32] := 0.60414171;
      W_o[5,33] := -0.01125434;
      W_o[5,34] := 0.53602260;
      W_o[5,35] := -0.02554985;
      W_o[5,36] := 0.12134581;
      W_o[5,37] := 0.08130677;
      W_o[5,38] := 0.47601295;
      W_o[5,39] := 0.06184123;
      W_o[6,0] := 0.43823916;
      W_o[6,1] := 0.04886893;
      W_o[6,2] := -0.72115153;
      W_o[6,3] := 0.53366846;
      W_o[6,4] := 0.14352611;
      W_o[6,5] := 0.27358714;
      W_o[6,6] := 1.15282750;
      W_o[6,7] := -0.53734303;
      W_o[6,8] := 0.10214026;
      W_o[6,9] := -0.33118525;
      W_o[6,10] := -0.18716197;
      W_o[6,11] := -0.26455408;
      W_o[6,12] := 0.97825962;
      W_o[6,13] := -0.17156628;
      W_o[6,14] := 0.04079279;
      W_o[6,15] := 0.20992042;
      W_o[6,16] := 0.19266997;
      W_o[6,17] := 0.39474788;
      W_o[6,18] := 0.49487942;
      W_o[6,19] := -0.59450352;
      W_o[6,20] := -0.62723535;
      W_o[6,21] := 0.23260640;
      W_o[6,22] := 0.70428210;
      W_o[6,23] := -0.57052928;
      W_o[6,24] := 2.01163483;
      W_o[6,25] := 1.53812528;
      W_o[6,26] := 0.15832324;
      W_o[6,27] := 0.01666135;
      W_o[6,28] := 0.11040143;
      W_o[6,29] := -0.30796206;
      W_o[6,30] := 0.70330209;
      W_o[6,31] := -0.19498926;
      W_o[6,32] := 0.43675256;
      W_o[6,33] := 0.28311005;
      W_o[6,34] := 2.10955501;
      W_o[6,35] := 0.06300426;
      W_o[6,36] := -0.06612100;
      W_o[6,37] := 0.24456324;
      W_o[6,38] := -0.06307534;
      W_o[6,39] := 0.85805798;
      W_o[7,0] := 0.03769494;
      W_o[7,1] := -0.15187448;
      W_o[7,2] := 0.09144486;
      W_o[7,3] := -0.05727371;
      W_o[7,4] := -0.34142601;
      W_o[7,5] := 0.31231621;
      W_o[7,6] := 0.12201753;
      W_o[7,7] := 0.15807615;
      W_o[7,8] := -0.11040714;
      W_o[7,9] := 0.17000853;
      W_o[7,10] := -0.22697128;
      W_o[7,11] := -0.60809618;
      W_o[7,12] := 0.17215836;
      W_o[7,13] := 0.31761804;
      W_o[7,14] := -0.22737864;
      W_o[7,15] := -0.11717512;
      W_o[7,16] := -0.05302644;
      W_o[7,17] := 0.26554984;
      W_o[7,18] := 0.28250584;
      W_o[7,19] := -0.15436935;
      W_o[7,20] := -0.33286601;
      W_o[7,21] := 0.64675540;
      W_o[7,22] := 0.03529684;
      W_o[7,23] := -0.64769369;
      W_o[7,24] := 1.23941433;
      W_o[7,25] := 1.17761362;
      W_o[7,26] := -0.46222582;
      W_o[7,27] := -0.28689626;
      W_o[7,28] := -0.04274225;
      W_o[7,29] := -0.00007054;
      W_o[7,30] := 0.25097835;
      W_o[7,31] := 0.01418501;
      W_o[7,32] := -0.11657754;
      W_o[7,33] := -0.23358633;
      W_o[7,34] := 0.18734637;
      W_o[7,35] := 0.05749683;
      W_o[7,36] := 0.03162088;
      W_o[7,37] := -0.04975284;
      W_o[7,38] := 0.03415622;
      W_o[7,39] := 0.03477194;
      R_i[0,0] := -0.11208162;
      R_i[0,1] := 0.02549788;
      R_i[0,2] := -0.17505924;
      R_i[0,3] := 0.19376156;
      R_i[0,4] := 0.16806792;
      R_i[0,5] := 0.17310023;
      R_i[0,6] := 0.23392540;
      R_i[0,7] := 0.24772970;
      R_i[1,0] := 0.12065984;
      R_i[1,1] := 1.14590645;
      R_i[1,2] := -0.48901820;
      R_i[1,3] := -0.41509745;
      R_i[1,4] := 0.09293488;
      R_i[1,5] := -0.53292608;
      R_i[1,6] := -0.76551837;
      R_i[1,7] := -1.31336629;
      R_i[2,0] := 0.30843908;
      R_i[2,1] := -0.34104937;
      R_i[2,2] := -1.87641382;
      R_i[2,3] := 0.96694976;
      R_i[2,4] := 0.27465352;
      R_i[2,5] := 0.13348614;
      R_i[2,6] := 0.10925449;
      R_i[2,7] := -0.03969188;
      R_i[3,0] := -0.47838771;
      R_i[3,1] := 0.29797852;
      R_i[3,2] := 0.66435951;
      R_i[3,3] := -4.26649761;
      R_i[3,4] := 0.10325183;
      R_i[3,5] := 1.01772487;
      R_i[3,6] := 0.25374600;
      R_i[3,7] := 0.20464782;
      R_i[4,0] := 0.32500589;
      R_i[4,1] := -0.23339252;
      R_i[4,2] := -0.22042707;
      R_i[4,3] := -0.07049563;
      R_i[4,4] := 1.06850040;
      R_i[4,5] := 0.45862436;
      R_i[4,6] := 0.19048849;
      R_i[4,7] := -0.10697714;
      R_i[5,0] := -0.13056895;
      R_i[5,1] := 0.09133054;
      R_i[5,2] := 0.12539217;
      R_i[5,3] := 0.23405170;
      R_i[5,4] := 0.28365436;
      R_i[5,5] := -0.09378310;
      R_i[5,6] := -0.37532172;
      R_i[5,7] := 0.33743879;
      R_i[6,0] := 0.45951205;
      R_i[6,1] := 0.01363123;
      R_i[6,2] := -0.29162151;
      R_i[6,3] := -0.22440894;
      R_i[6,4] := 0.06163742;
      R_i[6,5] := 0.38282368;
      R_i[6,6] := -0.96969271;
      R_i[6,7] := 0.10977434;
      R_i[7,0] := 0.20659432;
      R_i[7,1] := 0.27206531;
      R_i[7,2] := 0.59756833;
      R_i[7,3] := -0.40106091;
      R_i[7,4] := 0.29019260;
      R_i[7,5] := -0.57013249;
      R_i[7,6] := -0.22086233;
      R_i[7,7] := -1.44804525;
      R_f[0,0] := -0.90080142;
      R_f[0,1] := 0.76200789;
      R_f[0,2] := 0.75396901;
      R_f[0,3] := 0.18167311;
      R_f[0,4] := -0.70068061;
      R_f[0,5] := 0.19871995;
      R_f[0,6] := 0.67942381;
      R_f[0,7] := -1.24062347;
      R_f[1,0] := 0.60113764;
      R_f[1,1] := 0.83158749;
      R_f[1,2] := 0.45598811;
      R_f[1,3] := -0.72980219;
      R_f[1,4] := -0.50690895;
      R_f[1,5] := 0.34250832;
      R_f[1,6] := 0.19692127;
      R_f[1,7] := 0.53757608;
      R_f[2,0] := 0.36047983;
      R_f[2,1] := 0.07561547;
      R_f[2,2] := -1.04926670;
      R_f[2,3] := 0.20964669;
      R_f[2,4] := 0.65548646;
      R_f[2,5] := -0.14148460;
      R_f[2,6] := -0.28514028;
      R_f[2,7] := -0.50269139;
      R_f[3,0] := 0.28541896;
      R_f[3,1] := 0.81730789;
      R_f[3,2] := 1.12942076;
      R_f[3,3] := -1.25774288;
      R_f[3,4] := -0.45071271;
      R_f[3,5] := -0.27810058;
      R_f[3,6] := 0.34292591;
      R_f[3,7] := 0.19184071;
      R_f[4,0] := 0.30678338;
      R_f[4,1] := 0.29974887;
      R_f[4,2] := 0.06030706;
      R_f[4,3] := 0.09235083;
      R_f[4,4] := 1.58038485;
      R_f[4,5] := -0.05429833;
      R_f[4,6] := -0.01857536;
      R_f[4,7] := 0.17636755;
      R_f[5,0] := 0.90983230;
      R_f[5,1] := -0.17933325;
      R_f[5,2] := 0.50493723;
      R_f[5,3] := -1.05140698;
      R_f[5,4] := -0.31086558;
      R_f[5,5] := 0.52579153;
      R_f[5,6] := -0.87596011;
      R_f[5,7] := 1.19148707;
      R_f[6,0] := 0.74081868;
      R_f[6,1] := -0.65668273;
      R_f[6,2] := 0.54175776;
      R_f[6,3] := -1.03469229;
      R_f[6,4] := -0.06279287;
      R_f[6,5] := 0.25160038;
      R_f[6,6] := -0.27040246;
      R_f[6,7] := -0.19648477;
      R_f[7,0] := -0.22464477;
      R_f[7,1] := 0.34095991;
      R_f[7,2] := 1.24758875;
      R_f[7,3] := -0.71286923;
      R_f[7,4] := -0.48357251;
      R_f[7,5] := -0.06322154;
      R_f[7,6] := 0.18078713;
      R_f[7,7] := -0.41353473;
      R_g[0,0] := -2.33482742;
      R_g[0,1] := 0.26891232;
      R_g[0,2] := -0.62068361;
      R_g[0,3] := 1.05839896;
      R_g[0,4] := 0.97028506;
      R_g[0,5] := -0.01457710;
      R_g[0,6] := -0.11398745;
      R_g[0,7] := 0.24516355;
      R_g[1,0] := -0.11572418;
      R_g[1,1] := -2.35479641;
      R_g[1,2] := 0.09502196;
      R_g[1,3] := 0.01182066;
      R_g[1,4] := 0.12491781;
      R_g[1,5] := 0.00018514;
      R_g[1,6] := -0.13810089;
      R_g[1,7] := -0.12275805;
      R_g[2,0] := 0.10267565;
      R_g[2,1] := 0.09975577;
      R_g[2,2] := -1.91039574;
      R_g[2,3] := 0.88699478;
      R_g[2,4] := 0.83627421;
      R_g[2,5] := -0.05573991;
      R_g[2,6] := -0.02174967;
      R_g[2,7] := -0.06472150;
      R_g[3,0] := -0.03712863;
      R_g[3,1] := 0.03520567;
      R_g[3,2] := 0.00214308;
      R_g[3,3] := -1.63940406;
      R_g[3,4] := -0.30973291;
      R_g[3,5] := 0.00491419;
      R_g[3,6] := 0.05363122;
      R_g[3,7] := 0.04720224;
      R_g[4,0] := 0.02126839;
      R_g[4,1] := -0.05771927;
      R_g[4,2] := 0.66670042;
      R_g[4,3] := -0.78295749;
      R_g[4,4] := -2.66962981;
      R_g[4,5] := -0.05567581;
      R_g[4,6] := -0.03237662;
      R_g[4,7] := -0.01051190;
      R_g[5,0] := 0.17855854;
      R_g[5,1] := 0.28645414;
      R_g[5,2] := 0.40084702;
      R_g[5,3] := 1.08035278;
      R_g[5,4] := 0.47773901;
      R_g[5,5] := -2.19278741;
      R_g[5,6] := -0.20017563;
      R_g[5,7] := 0.14817512;
      R_g[6,0] := -0.16597822;
      R_g[6,1] := 0.06521239;
      R_g[6,2] := 0.30495486;
      R_g[6,3] := -0.52586186;
      R_g[6,4] := -0.41238609;
      R_g[6,5] := 0.18611307;
      R_g[6,6] := -1.59054327;
      R_g[6,7] := 0.01835538;
      R_g[7,0] := -0.12450181;
      R_g[7,1] := -0.22275996;
      R_g[7,2] := 0.13023397;
      R_g[7,3] := -0.52995551;
      R_g[7,4] := -0.57237208;
      R_g[7,5] := 0.16140953;
      R_g[7,6] := 0.00505236;
      R_g[7,7] := -2.26098657;
      R_o[0,0] := 1.05118394;
      R_o[0,1] := 1.61921883;
      R_o[0,2] := 0.40713361;
      R_o[0,3] := -0.12967324;
      R_o[0,4] := -0.75070161;
      R_o[0,5] := 0.60031158;
      R_o[0,6] := -0.96738613;
      R_o[0,7] := -0.49483040;
      R_o[1,0] := 0.40485424;
      R_o[1,1] := 0.52380055;
      R_o[1,2] := -0.32401261;
      R_o[1,3] := 0.06603508;
      R_o[1,4] := -0.39477521;
      R_o[1,5] := 0.40577486;
      R_o[1,6] := -0.40329638;
      R_o[1,7] := 0.24452984;
      R_o[2,0] := 0.32057163;
      R_o[2,1] := 0.76751244;
      R_o[2,2] := 3.85780931;
      R_o[2,3] := -0.80377811;
      R_o[2,4] := -0.76035577;
      R_o[2,5] := -0.06524058;
      R_o[2,6] := -0.31366009;
      R_o[2,7] := 0.89360225;
      R_o[3,0] := -0.04026479;
      R_o[3,1] := 0.06506599;
      R_o[3,2] := 0.94252461;
      R_o[3,3] := -1.12620234;
      R_o[3,4] := -1.53646183;
      R_o[3,5] := 0.08382892;
      R_o[3,6] := -0.13547981;
      R_o[3,7] := -0.12214545;
      R_o[4,0] := 0.35924345;
      R_o[4,1] := 0.13687599;
      R_o[4,2] := 0.84750414;
      R_o[4,3] := -0.98115104;
      R_o[4,4] := -1.33349466;
      R_o[4,5] := -0.73954433;
      R_o[4,6] := -0.11730482;
      R_o[4,7] := -0.01923019;
      R_o[5,0] := 0.71509749;
      R_o[5,1] := 2.16391206;
      R_o[5,2] := 1.45727324;
      R_o[5,3] := -0.44997519;
      R_o[5,4] := 0.08895559;
      R_o[5,5] := -0.45148489;
      R_o[5,6] := -0.91942245;
      R_o[5,7] := -0.81921595;
      R_o[6,0] := 0.77516019;
      R_o[6,1] := 0.79575026;
      R_o[6,2] := 0.57213145;
      R_o[6,3] := -0.32782549;
      R_o[6,4] := -1.04368973;
      R_o[6,5] := -0.26497081;
      R_o[6,6] := 0.46196660;
      R_o[6,7] := -0.07231894;
      R_o[7,0] := 0.64262104;
      R_o[7,1] := -0.09328733;
      R_o[7,2] := 0.49266991;
      R_o[7,3] := 0.05102121;
      R_o[7,4] := 0.01795285;
      R_o[7,5] := -0.13677078;
      R_o[7,6] := -0.15366967;
      R_o[7,7] := -0.31300050;
      B_i[0] := 0.47739047;
      B_i[1] := 1.16878533;
      B_i[2] := 0.07455011;
      B_i[3] := 0.71270287;
      B_i[4] := -0.25459385;
      B_i[5] := 0.41467166;
      B_i[6] := 1.58134580;
      B_i[7] := 0.48053345;
      B_f[0] := 1.96522069;
      B_f[1] := 2.15464544;
      B_f[2] := 0.96374005;
      B_f[3] := 3.17428517;
      B_f[4] := 1.05700183;
      B_f[5] := 2.83948231;
      B_f[6] := 1.68228626;
      B_f[7] := 2.85958314;
      B_g[0] := 0.84228754;
      B_g[1] := 0.67517793;
      B_g[2] := 1.40072227;
      B_g[3] := -0.51856840;
      B_g[4] := -1.00013328;
      B_g[5] := 0.12958716;
      B_g[6] := -0.54554117;
      B_g[7] := -0.30381307;
      B_o[0] := 3.60770607;
      B_o[1] := 1.64615154;
      B_o[2] := 2.89825439;
      B_o[3] := 2.80482626;
      B_o[4] := 2.26504564;
      B_o[5] := 3.94582796;
      B_o[6] := 3.44429064;
      B_o[7] := 2.25865412;
      FC_W[0,0] := -1.18992233;
      FC_W[0,1] := 0.05155103;
      FC_W[0,2] := -0.25555357;
      FC_W[0,3] := -1.68817246;
      FC_W[0,4] := 0.62249261;
      FC_W[0,5] := 2.72966671;
      FC_W[0,6] := 0.94766039;
      FC_W[0,7] := -0.05030653;
      FC_W[1,0] := 0.82415050;
      FC_W[1,1] := 0.10417762;
      FC_W[1,2] := 2.48935699;
      FC_W[1,3] := 0.90487832;
      FC_W[1,4] := -2.41745520;
      FC_W[1,5] := -2.44474673;
      FC_W[1,6] := -0.08907968;
      FC_W[1,7] := 0.45885682;
      FC_W[2,0] := -1.19081199;
      FC_W[2,1] := 0.06441317;
      FC_W[2,2] := -0.27430159;
      FC_W[2,3] := -1.68146050;
      FC_W[2,4] := 0.64268905;
      FC_W[2,5] := 2.70013452;
      FC_W[2,6] := 0.93640822;
      FC_W[2,7] := -0.06936958;
      FC_W[3,0] := -0.42120105;
      FC_W[3,1] := -0.03762053;
      FC_W[3,2] := -0.69488245;
      FC_W[3,3] := -2.14258838;
      FC_W[3,4] := 1.14586592;
      FC_W[3,5] := 1.54849517;
      FC_W[3,6] := -1.51691425;
      FC_W[3,7] := -0.79031748;
      FC_W[4,0] := -1.49379289;
      FC_W[4,1] := 0.29486084;
      FC_W[4,2] := -2.29751086;
      FC_W[4,3] := -1.71066320;
      FC_W[4,4] := -1.19953394;
      FC_W[4,5] := 0.04839557;
      FC_W[4,6] := 0.00004253;
      FC_W[4,7] := 1.18382549;
      FC_W[5,0] := -0.21551482;
      FC_W[5,1] := -1.39661205;
      FC_W[5,2] := 1.55288088;
      FC_W[5,3] := -0.20406686;
      FC_W[5,4] := 0.61307526;
      FC_W[5,5] := -1.18333137;
      FC_W[5,6] := 0.65153670;
      FC_W[5,7] := -0.30164590;
      FC_W[6,0] := 0.29921451;
      FC_W[6,1] := -2.77646971;
      FC_W[6,2] := 0.34926391;
      FC_W[6,3] := -1.64131200;
      FC_W[6,4] := 1.16665757;
      FC_W[6,5] := -0.32929334;
      FC_W[6,6] := 1.03012013;
      FC_W[6,7] := -1.66025639;
      FC_W[7,0] := -0.41906875;
      FC_W[7,1] := -0.05154445;
      FC_W[7,2] := -0.70114154;
      FC_W[7,3] := -2.15366507;
      FC_W[7,4] := 1.14648783;
      FC_W[7,5] := 1.57242584;
      FC_W[7,6] := -1.49940395;
      FC_W[7,7] := -0.77594888;
      FC_W[8,0] := -0.43902808;
      FC_W[8,1] := -0.03909670;
      FC_W[8,2] := -0.71527648;
      FC_W[8,3] := -2.07963490;
      FC_W[8,4] := 1.21875131;
      FC_W[8,5] := 1.52684188;
      FC_W[8,6] := -1.52031815;
      FC_W[8,7] := -0.76095748;
      FC_W[9,0] := -0.42732900;
      FC_W[9,1] := -0.03466158;
      FC_W[9,2] := -0.68948311;
      FC_W[9,3] := -2.14737368;
      FC_W[9,4] := 1.15473747;
      FC_W[9,5] := 1.56467116;
      FC_W[9,6] := -1.51235425;
      FC_W[9,7] := -0.78273284;
      FC_W[10,0] := -0.58327764;
      FC_W[10,1] := 1.46903265;
      FC_W[10,2] := -0.12583148;
      FC_W[10,3] := -0.77770352;
      FC_W[10,4] := 0.44943938;
      FC_W[10,5] := 1.18295085;
      FC_W[10,6] := -1.91800594;
      FC_W[10,7] := 0.32411379;
      FC_W[11,0] := 0.20698918;
      FC_W[11,1] := 1.86358893;
      FC_W[11,2] := -0.93361831;
      FC_W[11,3] := -1.29574013;
      FC_W[11,4] := -0.03512571;
      FC_W[11,5] := -0.29252213;
      FC_W[11,6] := 0.28302547;
      FC_W[11,7] := -1.40581882;
      FC_W[12,0] := 0.39387086;
      FC_W[12,1] := 1.50321007;
      FC_W[12,2] := -0.68883723;
      FC_W[12,3] := -1.38207150;
      FC_W[12,4] := 0.04493435;
      FC_W[12,5] := -0.39445713;
      FC_W[12,6] := -0.09016615;
      FC_W[12,7] := -1.20629704;
      FC_W[13,0] := -0.68904585;
      FC_W[13,1] := 0.38990816;
      FC_W[13,2] := 4.25386047;
      FC_W[13,3] := -1.10076106;
      FC_W[13,4] := -1.86902809;
      FC_W[13,5] := -0.19047922;
      FC_W[13,6] := 0.11304056;
      FC_W[13,7] := 0.72004426;
      FC_W[14,0] := -2.93907404;
      FC_W[14,1] := -1.89689541;
      FC_W[14,2] := -0.33583719;
      FC_W[14,3] := 0.87999964;
      FC_W[14,4] := -2.06177592;
      FC_W[14,5] := 0.70418972;
      FC_W[14,6] := -1.52928364;
      FC_W[14,7] := -2.70884418;
      FC_W[15,0] := -0.21864611;
      FC_W[15,1] := 1.95235348;
      FC_W[15,2] := -1.01023436;
      FC_W[15,3] := -1.06552947;
      FC_W[15,4] := -0.29395279;
      FC_W[15,5] := -0.18908904;
      FC_W[15,6] := 0.54388875;
      FC_W[15,7] := -1.83758295;
      FC_W[16,0] := -1.21153963;
      FC_W[16,1] := -3.00696540;
      FC_W[16,2] := 0.27524677;
      FC_W[16,3] := 0.12779871;
      FC_W[16,4] := -0.98358935;
      FC_W[16,5] := 0.55670607;
      FC_W[16,6] := -2.62852859;
      FC_W[16,7] := -0.72020465;
      FC_W[17,0] := 2.03641272;
      FC_W[17,1] := -2.40191722;
      FC_W[17,2] := 1.36396074;
      FC_W[17,3] := -0.75134295;
      FC_W[17,4] := 1.27749395;
      FC_W[17,5] := -0.64430392;
      FC_W[17,6] := -2.46128988;
      FC_W[17,7] := 2.50009131;
      FC_W[18,0] := 1.15559602;
      FC_W[18,1] := -0.17385845;
      FC_W[18,2] := -4.94069910;
      FC_W[18,3] := -0.70903516;
      FC_W[18,4] := -0.56411159;
      FC_W[18,5] := 1.44895744;
      FC_W[18,6] := 1.31446946;
      FC_W[18,7] := -0.49564546;
      FC_W[19,0] := 0.16732359;
      FC_W[19,1] := 1.55335963;
      FC_W[19,2] := 0.38663110;
      FC_W[19,3] := -1.15490484;
      FC_W[19,4] := 0.16659181;
      FC_W[19,5] := -0.77653676;
      FC_W[19,6] := -0.28400528;
      FC_W[19,7] := -1.09486878;
      FC_W[20,0] := -0.27414966;
      FC_W[20,1] := 2.61213183;
      FC_W[20,2] := -0.27200100;
      FC_W[20,3] := 0.60704172;
      FC_W[20,4] := -1.86421537;
      FC_W[20,5] := 0.47701240;
      FC_W[20,6] := -1.07750309;
      FC_W[20,7] := 1.48161185;
      FC_W[21,0] := 2.28589869;
      FC_W[21,1] := -1.45107174;
      FC_W[21,2] := -0.91967463;
      FC_W[21,3] := -0.98829103;
      FC_W[21,4] := -0.53788638;
      FC_W[21,5] := 1.15463293;
      FC_W[21,6] := 1.29627419;
      FC_W[21,7] := -2.03720641;
      FC_W[22,0] := 0.70766956;
      FC_W[22,1] := -0.16230604;
      FC_W[22,2] := 2.38536215;
      FC_W[22,3] := -3.18115830;
      FC_W[22,4] := -4.12445784;
      FC_W[22,5] := 0.27941021;
      FC_W[22,6] := -0.13647506;
      FC_W[22,7] := -0.44242245;
      FC_W[23,0] := -1.06704283;
      FC_W[23,1] := 0.64061731;
      FC_W[23,2] := 4.17096949;
      FC_W[23,3] := -1.59397840;
      FC_W[23,4] := -1.34815049;
      FC_W[23,5] := 0.38533959;
      FC_W[23,6] := -0.84740913;
      FC_W[23,7] := 0.35435632;
      FC_W[24,0] := 0.79453409;
      FC_W[24,1] := -0.20100924;
      FC_W[24,2] := 2.19239259;
      FC_W[24,3] := -3.21025372;
      FC_W[24,4] := -4.16017342;
      FC_W[24,5] := 0.32382092;
      FC_W[24,6] := -0.05922369;
      FC_W[24,7] := -0.48731399;
      FC_W[25,0] := 0.79488528;
      FC_W[25,1] := -0.20141180;
      FC_W[25,2] := 2.20286703;
      FC_W[25,3] := -3.21136475;
      FC_W[25,4] := -4.16547203;
      FC_W[25,5] := 0.32160446;
      FC_W[25,6] := -0.06135242;
      FC_W[25,7] := -0.48731378;
      FC_W[26,0] := -1.22062659;
      FC_W[26,1] := 0.45275605;
      FC_W[26,2] := 3.50765562;
      FC_W[26,3] := -1.81133246;
      FC_W[26,4] := -2.32191133;
      FC_W[26,5] := -0.85800213;
      FC_W[26,6] := -1.03187132;
      FC_W[26,7] := 0.84669930;
      FC_W[27,0] := 2.16321373;
      FC_W[27,1] := -1.26625168;
      FC_W[27,2] := -1.54215634;
      FC_W[27,3] := -0.51378232;
      FC_W[27,4] := -0.03297012;
      FC_W[27,5] := 1.24442351;
      FC_W[27,6] := 1.31537867;
      FC_W[27,7] := -1.86622298;
      FC_W[28,0] := -1.85206807;
      FC_W[28,1] := -1.12244534;
      FC_W[28,2] := -1.02892709;
      FC_W[28,3] := -2.12493491;
      FC_W[28,4] := 0.42766815;
      FC_W[28,5] := -0.43299294;
      FC_W[28,6] := 0.84881854;
      FC_W[28,7] := 0.19362010;
      FC_W[29,0] := -0.72036493;
      FC_W[29,1] := 0.19177595;
      FC_W[29,2] := -2.20158601;
      FC_W[29,3] := 3.11478376;
      FC_W[29,4] := 3.95264387;
      FC_W[29,5] := -0.30077153;
      FC_W[29,6] := 0.08013711;
      FC_W[29,7] := 0.48923638;
      FC_W[30,0] := 0.70360428;
      FC_W[30,1] := -0.15897189;
      FC_W[30,2] := 2.38808751;
      FC_W[30,3] := -3.17935729;
      FC_W[30,4] := -4.12390041;
      FC_W[30,5] := 0.27836224;
      FC_W[30,6] := -0.13839228;
      FC_W[30,7] := -0.43985024;
      FC_W[31,0] := 0.66204989;
      FC_W[31,1] := -0.15782984;
      FC_W[31,2] := 2.41914916;
      FC_W[31,3] := -3.15487289;
      FC_W[31,4] := -4.07718945;
      FC_W[31,5] := 0.25418258;
      FC_W[31,6] := -0.15442266;
      FC_W[31,7] := -0.42680934;
      FC_W[32,0] := 0.79047048;
      FC_W[32,1] := -0.23469672;
      FC_W[32,2] := 2.29716516;
      FC_W[32,3] := -3.24202681;
      FC_W[32,4] := -4.15815735;
      FC_W[32,5] := 0.30668151;
      FC_W[32,6] := -0.05686283;
      FC_W[32,7] := -0.50771844;
      FC_W[33,0] := 0.75455624;
      FC_W[33,1] := -0.25742382;
      FC_W[33,2] := 2.35943079;
      FC_W[33,3] := -3.22433543;
      FC_W[33,4] := -4.10108995;
      FC_W[33,5] := 0.25491622;
      FC_W[33,6] := -0.07580780;
      FC_W[33,7] := -0.49778089;
      FC_W[34,0] := 0.71609271;
      FC_W[34,1] := -0.21596618;
      FC_W[34,2] := 2.39747453;
      FC_W[34,3] := -3.21923876;
      FC_W[34,4] := -4.10705996;
      FC_W[34,5] := 0.26319802;
      FC_W[34,6] := -0.10984568;
      FC_W[34,7] := -0.47146788;
      FC_W[35,0] := 0.82340604;
      FC_W[35,1] := -0.23696223;
      FC_W[35,2] := 2.22725129;
      FC_W[35,3] := -3.24754643;
      FC_W[35,4] := -4.16000032;
      FC_W[35,5] := 0.35599440;
      FC_W[35,6] := -0.02254982;
      FC_W[35,7] := -0.52403253;
      FC_W[36,0] := 1.70248604;
      FC_W[36,1] := 0.11325528;
      FC_W[36,2] := -0.55486101;
      FC_W[36,3] := -1.79293418;
      FC_W[36,4] := -3.01944804;
      FC_W[36,5] := 1.24814284;
      FC_W[36,6] := 0.53546667;
      FC_W[36,7] := -0.78272438;
      FC_W[37,0] := 0.84245664;
      FC_W[37,1] := -0.24852155;
      FC_W[37,2] := 2.21305323;
      FC_W[37,3] := -3.24593639;
      FC_W[37,4] := -4.15289927;
      FC_W[37,5] := 0.36589786;
      FC_W[37,6] := -0.00642151;
      FC_W[37,7] := -0.53890944;
      FC_W[38,0] := -2.70351076;
      FC_W[38,1] := -2.30757785;
      FC_W[38,2] := -0.31027862;
      FC_W[38,3] := 0.69808859;
      FC_W[38,4] := -1.93468404;
      FC_W[38,5] := 0.86156154;
      FC_W[38,6] := -1.85448647;
      FC_W[38,7] := -2.37202263;
      FC_W[39,0] := -3.07146120;
      FC_W[39,1] := -2.31486058;
      FC_W[39,2] := -0.36967734;
      FC_W[39,3] := 0.85301226;
      FC_W[39,4] := -2.18805957;
      FC_W[39,5] := 0.90125442;
      FC_W[39,6] := -1.85495472;
      FC_W[39,7] := -2.75822377;
      FC_B[0] := -0.13849375;
      FC_B[1] := -0.99999899;
      FC_B[2] := -0.13808991;
      FC_B[3] := -0.50583917;
      FC_B[4] := -0.07021909;
      FC_B[5] := -0.04431012;
      FC_B[6] := 0.21439837;
      FC_B[7] := -0.49694595;
      FC_B[8] := -0.46466905;
      FC_B[9] := -0.50298262;
      FC_B[10] := -0.66974354;
      FC_B[11] := -0.89998204;
      FC_B[12] := -0.93942428;
      FC_B[13] := -1.98418629;
      FC_B[14] := 0.76125818;
      FC_B[15] := -0.80674237;
      FC_B[16] := 0.61973643;
      FC_B[17] := -0.10940201;
      FC_B[18] := 1.23516512;
      FC_B[19] := -1.18503582;
      FC_B[20] := -0.73241270;
      FC_B[21] := 0.09495984;
      FC_B[22] := -2.61826062;
      FC_B[23] := -2.19209623;
      FC_B[24] := -2.57054734;
      FC_B[25] := -2.57508588;
      FC_B[26] := -2.22407436;
      FC_B[27] := 0.50726670;
      FC_B[28] := 0.10793630;
      FC_B[29] := 2.51168299;
      FC_B[30] := -2.61885405;
      FC_B[31] := -2.61374116;
      FC_B[32] := -2.60812306;
      FC_B[33] := -2.60557532;
      FC_B[34] := -2.62382841;
      FC_B[35] := -2.59056973;
      FC_B[36] := -1.10703635;
      FC_B[37] := -2.58282399;
      FC_B[38] := 0.78152573;
      FC_B[39] := 0.85155326;

END_DATA_BLOCK
